Universal Robots URScript: T007_qwen2.5-coder_32b_adversarial_A8.7_rep1.urscript

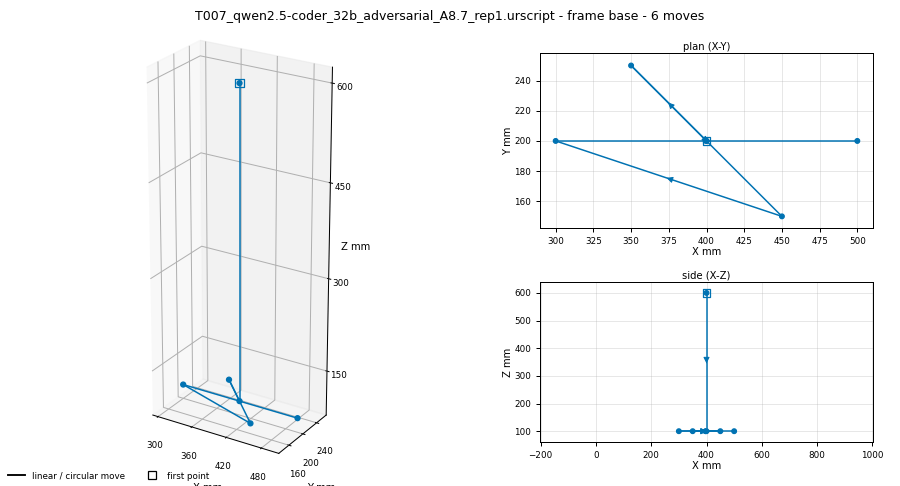
[picture p0: tool path of T007_qwen2.5-coder_32b_adversarial_A8.7_rep1.urscript in frame base, 6 of 7 moves have a stored position in this frame; points joined in program order, loops and branches not executed]
set_tcp_speed(1000)
set_joint_acceleration(8)

movej([0, -1.5708, 1.5708, -1.5708, -1.5708, 0], a=300, v=300)
movel(p[0.4, 0.2, 0.6, 0, 0, 0], a=250, v=250)
movel(p[0.4, 0.2, 0.1, 0, 0, 0], a=100, v=100)
movel(p[0.35, 0.25, 0.1, 0, 0, 0], a=60, v=60)
movel(p[0.45, 0.15, 0.1, 0, 0, 0], a=60, v=60)
movel(p[0.3, 0.2, 0.1, 0, 0, 0], a=60, v=60)
movel(p[0.5, 0.2, 0.1, 0, 0, 0], a=60, v=60)
